(* IEC 61131-3 sources: trust-platform/tests/corpus, 4 files *)

(* ---- control_flow.st ---- *)
(* Test corpus: Control flow statements *)

PROGRAM TestControlFlow

VAR
    i, j, k : INT;
    condition : BOOL;
    state : INT;
    result : INT;
    sum : INT;
    arr : ARRAY[0..9] OF INT;
END_VAR

(* Simple IF *)
IF condition THEN
    result := 1;
END_IF

(* IF-ELSE *)
IF condition THEN
    result := 1;
ELSE
    result := 0;
END_IF

(* IF-ELSIF-ELSE *)
IF i < 0 THEN
    result := -1;
ELSIF i = 0 THEN
    result := 0;
ELSIF i > 0 AND i < 10 THEN
    result := 1;
ELSE
    result := 2;
END_IF

(* Nested IF *)
IF condition THEN
    IF i > 0 THEN
        result := 1;
    ELSE
        result := 2;
    END_IF
END_IF

(* Simple CASE *)
CASE state OF
    0: result := 0;
    1: result := 1;
    2: result := 2;
END_CASE

(* CASE with multiple labels *)
CASE state OF
    0, 1, 2:
        result := 0;
    3, 4, 5:
        result := 1;
    6..10:
        result := 2;
END_CASE

(* CASE with ELSE *)
CASE state OF
    0:
        result := 0;
    1:
        result := 1;
ELSE
    result := -1;
END_CASE

(* CASE with multiple statements *)
CASE state OF
    0:
        result := 0;
        condition := FALSE;
    1:
        result := 1;
        condition := TRUE;
END_CASE

(* Simple FOR *)
FOR i := 0 TO 9 DO
    arr[i] := i;
END_FOR

(* FOR with BY *)
FOR i := 0 TO 100 BY 10 DO
    sum := sum + i;
END_FOR

(* FOR counting down *)
FOR i := 10 TO 0 BY -1 DO
    arr[i] := i * 2;
END_FOR

(* Nested FOR *)
FOR i := 0 TO 9 DO
    FOR j := 0 TO 9 DO
        result := i * 10 + j;
    END_FOR
END_FOR

(* Simple WHILE *)
i := 0;
WHILE i < 10 DO
    sum := sum + i;
    i := i + 1;
END_WHILE

(* WHILE with complex condition *)
WHILE i < 10 AND NOT condition DO
    i := i + 1;
END_WHILE

(* Nested WHILE *)
i := 0;
WHILE i < 5 DO
    j := 0;
    WHILE j < 5 DO
        result := i * j;
        j := j + 1;
    END_WHILE
    i := i + 1;
END_WHILE

(* Simple REPEAT *)
i := 0;
REPEAT
    sum := sum + i;
    i := i + 1;
UNTIL i >= 10
END_REPEAT

(* REPEAT with complex condition *)
REPEAT
    i := i + 1;
    condition := i MOD 2 = 0;
UNTIL condition OR i > 100
END_REPEAT

(* EXIT from loop *)
FOR i := 0 TO 100 DO
    IF i > 50 THEN
        EXIT;
    END_IF
    sum := sum + i;
END_FOR

(* CONTINUE in loop *)
FOR i := 0 TO 9 DO
    IF i MOD 2 = 0 THEN
        CONTINUE;
    END_IF
    sum := sum + i;
END_FOR

(* EXIT from nested loop *)
FOR i := 0 TO 9 DO
    FOR j := 0 TO 9 DO
        IF i * j > 50 THEN
            EXIT;
        END_IF
    END_FOR
END_FOR

(* Empty statement *)
;

(* Multiple empty statements *)
;;

END_PROGRAM

(* Function with RETURN *)
FUNCTION CalcSum : INT
VAR_INPUT
    n : INT;
END_VAR
VAR
    i : INT;
    sum : INT;
END_VAR

IF n <= 0 THEN
    RETURN;
END_IF

FOR i := 1 TO n DO
    sum := sum + i;
END_FOR

CalcSum := sum;
END_FUNCTION

(* Function with early RETURN *)
FUNCTION FindIndex : INT
VAR_INPUT
    arr : ARRAY[0..9] OF INT;
    value : INT;
END_VAR
VAR
    i : INT;
END_VAR

FOR i := 0 TO 9 DO
    IF arr[i] = value THEN
        FindIndex := i;
        RETURN;
    END_IF
END_FOR

FindIndex := -1;
END_FUNCTION

(* Complex control flow *)
FUNCTION_BLOCK FB_StateMachine
VAR
    state : INT;
    counter : INT;
    done : BOOL;
END_VAR

CASE state OF
    0: (* Init *)
        counter := 0;
        state := 1;

    1: (* Process *)
        WHILE counter < 100 AND NOT done DO
            counter := counter + 1;
            IF counter MOD 10 = 0 THEN
                (* Check condition *)
                IF counter > 50 THEN
                    done := TRUE;
                    EXIT;
                END_IF
            END_IF
        END_WHILE

        IF done THEN
            state := 2;
        END_IF

    2: (* Done *)
        ; (* Empty - wait *)
END_CASE

END_FUNCTION_BLOCK

(* ---- declarations.st ---- *)
(* Test corpus: Variable declarations and modifiers *)

PROGRAM TestDeclarations

(* Basic variable block *)
VAR
    simpleVar : INT;
    multipleVars, anotherVar : BOOL;
    initialized : REAL := 3.14;
END_VAR

(* Input variables *)
VAR_INPUT
    inputBool : BOOL;
    inputInt : INT := 100;
END_VAR

(* Output variables *)
VAR_OUTPUT
    outputStatus : BOOL;
    outputValue : REAL;
END_VAR

(* In-out variables *)
VAR_IN_OUT
    inoutData : ARRAY[0..9] OF INT;
END_VAR

(* Temporary variables *)
VAR_TEMP
    tempCounter : INT;
    tempBuffer : STRING[80];
END_VAR

(* Constant variables *)
VAR CONSTANT
    PI : REAL := 3.14159;
    MAX_SIZE : INT := 1000;
END_VAR

(* Retain variables *)
VAR RETAIN
    persistentCounter : UDINT;
END_VAR

(* Non-retain variables *)
VAR NON_RETAIN
    volatileData : REAL;
END_VAR

(* Persistent variables *)
VAR PERSISTENT
    savedState : INT;
END_VAR

(* All elementary types *)
VAR
    boolVal : BOOL;
    sintVal : SINT;
    intVal : INT;
    dintVal : DINT;
    lintVal : LINT;
    usintVal : USINT;
    uintVal : UINT;
    udintVal : UDINT;
    ulintVal : ULINT;
    realVal : REAL;
    lrealVal : LREAL;
    byteVal : BYTE;
    wordVal : WORD;
    dwordVal : DWORD;
    lwordVal : LWORD;
    stringVal : STRING;
    stringFixed : STRING[100];
    wstringVal : WSTRING;
    timeVal : TIME;
    ltimeVal : LTIME;
    dateVal : DATE;
    todVal : TIME_OF_DAY;
    dtVal : DATE_AND_TIME;
END_VAR

END_PROGRAM

(* Global variables - must be in CONFIGURATION per IEC 61131-3 *)
CONFIGURATION GlobalConfig
VAR_GLOBAL
    GlobalCounter : UDINT;
    GlobalStatus : BOOL;
END_VAR

VAR_GLOBAL CONSTANT
    APP_VERSION : STRING := '1.0.0';
END_VAR
END_CONFIGURATION

(* External variables *)
PROGRAM TestExternal
VAR_EXTERNAL
    ExternalRef : REAL;
END_VAR
END_PROGRAM

(* Static variables in function block *)
FUNCTION_BLOCK FB_WithStatic
VAR_STAT
    callCount : UDINT;
END_VAR

callCount := callCount + 1;
END_FUNCTION_BLOCK

(* Type declarations *)
TYPE MyInt : INT; END_TYPE

TYPE MyRange : INT (0..100); END_TYPE

TYPE MyArray : ARRAY[0..9] OF INT; END_TYPE

TYPE MyArray2D : ARRAY[0..9, 0..9] OF REAL; END_TYPE

TYPE MyPointer : POINTER TO INT; END_TYPE

TYPE MyRef : REF_TO REAL; END_TYPE

TYPE MyString : STRING[255]; END_TYPE

TYPE MyStruct :
STRUCT
    field1 : INT;
    field2 : REAL;
    field3 : STRING[50];
END_STRUCT
END_TYPE

TYPE MyUnion :
UNION
    asInt : DINT;
    asReal : REAL;
    asBytes : ARRAY[0..3] OF BYTE;
END_UNION
END_TYPE

TYPE Color :
(
    Red := 0,
    Green := 1,
    Blue := 2
);
END_TYPE

(* Function with parameters *)
FUNCTION Add : INT
VAR_INPUT
    a : INT;
    b : INT;
END_VAR

Add := a + b;
END_FUNCTION

(* Function block with inheritance *)
FUNCTION_BLOCK FB_Child EXTENDS FB_Parent IMPLEMENTS I_Interface
VAR
    childVar : INT;
END_VAR
END_FUNCTION_BLOCK

(* Interface declaration *)
INTERFACE I_Counter
    METHOD Increment : INT
    END_METHOD

    METHOD Reset
    END_METHOD

    PROPERTY Count : INT
    END_PROPERTY
END_INTERFACE

(* Method with access modifiers *)
FUNCTION_BLOCK FB_AccessTest
VAR PUBLIC
    publicVar : INT;
END_VAR

VAR PRIVATE
    privateVar : INT;
END_VAR

PROTECTED METHOD ProtectedMethod
END_METHOD

PUBLIC METHOD PublicMethod
END_METHOD

PRIVATE METHOD PrivateMethod
END_METHOD
END_FUNCTION_BLOCK

(* Property with getter and setter *)
FUNCTION_BLOCK FB_PropertyTest
VAR
    _value : INT;
END_VAR

PROPERTY Value : INT
    GET
        Value := _value;
    END_GET
    SET
        _value := Value;
    END_SET
END_PROPERTY
END_FUNCTION_BLOCK

(* Namespace *)
NAMESPACE MyApp
    FUNCTION_BLOCK FB_Nested
    END_FUNCTION_BLOCK
END_NAMESPACE

(* ---- expressions.st ---- *)
(* Test corpus: Expressions and operator precedence *)

PROGRAM TestExpressions

VAR
    a, b, c, d : INT;
    x, y, z : REAL;
    p, q, r : BOOL;
    s1, s2 : STRING;
    arr : ARRAY[0..9] OF INT;
    ptr : POINTER TO INT;
    fb : FB_Test;
END_VAR

(* ============================================= *)
(* Arithmetic operators *)
(* ============================================= *)

(* Addition *)
a := 1 + 2;
a := b + c;
x := 1.0 + 2.5;

(* Subtraction *)
a := 5 - 3;
a := b - c;
x := 10.0 - 3.5;

(* Multiplication *)
a := 3 * 4;
a := b * c;
x := 2.0 * 3.14;

(* Division *)
a := 10 / 2;
x := 10.0 / 3.0;

(* Modulo *)
a := 10 MOD 3;
a := b MOD c;

(* Exponentiation - right associative *)
x := 2.0 ** 3.0;
x := 2.0 ** 3.0 ** 2.0;  (* = 2^(3^2) = 2^9 = 512 *)

(* Unary operators *)
a := -b;
a := +c;
x := -3.14;

(* ============================================= *)
(* Comparison operators *)
(* ============================================= *)

p := a = b;
p := a <> b;
p := a < b;
p := a <= b;
p := a > b;
p := a >= b;

(* String comparison *)
p := s1 = s2;
p := s1 < s2;

(* ============================================= *)
(* Logical operators *)
(* ============================================= *)

(* AND *)
p := q AND r;
p := q & r;

(* OR *)
p := q OR r;

(* XOR *)
p := q XOR r;

(* NOT *)
p := NOT q;

(* ============================================= *)
(* Bitwise operators *)
(* ============================================= *)

a := b AND c;
a := b OR c;
a := b XOR c;
a := NOT b;

(* ============================================= *)
(* Operator precedence tests *)
(* ============================================= *)

(* Precedence: * before + *)
a := 1 + 2 * 3;         (* = 1 + 6 = 7 *)
a := (1 + 2) * 3;       (* = 3 * 3 = 9 *)

(* Precedence: AND before OR *)
p := TRUE OR FALSE AND FALSE;     (* = TRUE OR FALSE = TRUE *)
p := (TRUE OR FALSE) AND FALSE;   (* = TRUE AND FALSE = FALSE *)

(* Precedence: comparison before logical *)
p := a < b AND c > d;   (* = (a < b) AND (c > d) *)

(* Precedence: arithmetic before comparison *)
p := a + b < c + d;     (* = (a + b) < (c + d) *)

(* Precedence: NOT has highest priority *)
p := NOT q AND r;       (* = (NOT q) AND r *)
p := NOT (q AND r);     (* = NOT (q AND r) *)

(* Complex precedence *)
a := 1 + 2 * 3 - 4 / 2;     (* = 1 + 6 - 2 = 5 *)
p := a > b OR c < d AND NOT r;  (* = (a > b) OR ((c < d) AND (NOT r)) *)

(* Power is right associative *)
x := 2.0 ** 2.0 ** 3.0;     (* = 2^(2^3) = 2^8 = 256 *)

(* ============================================= *)
(* Parenthesized expressions *)
(* ============================================= *)

a := (b);
a := ((b));
a := (b + c);
a := (b + c) * d;
a := ((b + c) * (d - a));

(* ============================================= *)
(* Function calls *)
(* ============================================= *)

x := SIN(3.14);
x := ABS(-42);
a := MAX(b, c);
x := SQRT(y);

(* Nested function calls *)
x := SIN(COS(3.14));
x := ABS(MIN(a, b));

(* Function call in expression *)
x := 2.0 * SIN(y) + 1.0;

(* Named parameters *)
(* result := MyFunc(param1 := 10, param2 := 20); *)

(* ============================================= *)
(* Array indexing *)
(* ============================================= *)

a := arr[0];
a := arr[b];
a := arr[b + 1];
a := arr[b * 2 + c];

(* Multi-dimensional *)
(* a := matrix[i, j]; *)
(* a := matrix[i][j]; *)

(* ============================================= *)
(* Field access *)
(* ============================================= *)

a := fb.value;
x := fb.data.x;
a := fb.nested.deep.value;

(* Method call *)
a := fb.GetValue();
fb.SetValue(10);

(* ============================================= *)
(* Pointer operations *)
(* ============================================= *)

(* Dereference *)
a := ptr^;

(* Address-of *)
ptr := ADR(a);

(* SIZEOF *)
a := SIZEOF(INT);
a := SIZEOF(arr);
a := SIZEOF(fb);

(* ============================================= *)
(* Special expressions *)
(* ============================================= *)

(* THIS and SUPER *)
(* a := THIS.value; *)
(* a := SUPER.GetValue(); *)

(* Direct addresses *)
(* a := %IW10; *)
(* p := %IX0.0; *)

(* Typed literals in expressions *)
a := INT#42 + INT#10;
x := REAL#3.14 * REAL#2.0;

(* ============================================= *)
(* Complex expressions *)
(* ============================================= *)

(* Combined arithmetic and logic *)
p := (a + b > c) AND (d - a < 10) OR NOT q;

(* Expression with function call and array *)
a := arr[MAX(b, c)] + ABS(d);

(* Expression with field access *)
x := fb.value * SIN(fb.angle);

(* Very complex expression *)
x := ((a + b) * SIN(c / d)) / (SQRT(y ** 2.0 + z ** 2.0) + 1.0);

END_PROGRAM

(* Function block for testing *)
FUNCTION_BLOCK FB_Test
VAR
    value : INT;
    angle : REAL;
    data : ST_Data;
    nested : FB_Nested;
END_VAR

METHOD GetValue : INT
    GetValue := value;
END_METHOD

METHOD SetValue
VAR_INPUT
    newValue : INT;
END_VAR
    value := newValue;
END_METHOD
END_FUNCTION_BLOCK

FUNCTION_BLOCK FB_Nested
VAR
    deep : ST_Deep;
END_VAR
END_FUNCTION_BLOCK

TYPE ST_Data :
STRUCT
    x : REAL;
    y : REAL;
END_STRUCT
END_TYPE

TYPE ST_Deep :
STRUCT
    value : INT;
END_STRUCT
END_TYPE

(* Test expression edge cases *)
FUNCTION TestEdgeCases : BOOL
VAR
    a : INT;
    x : REAL;
    p : BOOL;
END_VAR

(* Double negation *)
a := --5;
a := -(-a);
x := --3.14;

(* NOT NOT *)
p := NOT NOT TRUE;
p := NOT NOT p;

(* Chained comparisons need explicit grouping *)
p := (a < 5) AND (5 < 10);

(* Very deep nesting *)
a := ((((((1 + 2) * 3) - 4) / 5) MOD 6) + 7);

TestEdgeCases := TRUE;
END_FUNCTION

(* ---- literals.st ---- *)
(* Test corpus: All literal types *)

PROGRAM TestLiterals

VAR
    (* Integer literals *)
    intDec : INT := 123;
    intNeg : INT := -456;
    intZero : INT := 0;
    intWithUnder : DINT := 1_000_000;

    (* Hexadecimal literals *)
    intHex : DWORD := 16#FF;
    intHexLower : DWORD := 16#ff;
    intHexMixed : DWORD := 16#DeAdBeEf;
    intHexUnder : DWORD := 16#DEAD_BEEF;

    (* Binary literals *)
    intBin : BYTE := 2#10101010;
    intBinUnder : WORD := 2#1111_0000_1111_0000;

    (* Octal literals *)
    intOct : INT := 8#77;
    intOctUnder : INT := 8#7_7_7;

    (* Real literals *)
    realSimple : REAL := 3.14;
    realNeg : REAL := -2.718;
    realZero : REAL := 0.0;
    realSmall : REAL := 0.001;
    realWithUnder : LREAL := 1_000.000_001;

    (* Scientific notation *)
    realSci1 : LREAL := 1.0E10;
    realSci2 : LREAL := 2.5e-3;
    realSci3 : LREAL := 6.022E+23;
    realSciNeg : LREAL := -1.6E-19;

    (* Boolean literals *)
    boolTrue : BOOL := TRUE;
    boolFalse : BOOL := FALSE;
    boolTrueLower : BOOL := true;
    boolFalseLower : BOOL := false;

    (* String literals - single quote *)
    strEmpty : STRING := '';
    strSimple : STRING := 'Hello, World!';
    strWithEscape : STRING := 'Line1$NLine2';
    strWithQuote : STRING := 'It$'s working';
    strPath : STRING := 'C:\Program Files\App';

    (* Wide string literals - double quote *)
    wstrEmpty : WSTRING := "";
    wstrSimple : WSTRING := "Wide string";
    wstrUnicode : WSTRING := "日本語";

    (* Time literals *)
    timeSimple : TIME := T#1s;
    timeLong : TIME := TIME#1h30m45s;
    timeMs : TIME := T#100ms;
    timeComplex : TIME := T#1d2h3m4s5ms;
    timeUnder : TIME := T#1000ms;
    ltimeVal : LTIME := LTIME#1h;

    (* Date literals *)
    dateSimple : DATE := D#2024-01-15;
    dateFull : DATE := DATE#2024-12-31;

    (* Time of day literals *)
    todSimple : TIME_OF_DAY := TOD#12:30:00;
    todFull : TIME_OF_DAY := TIME_OF_DAY#23:59:59.999;
    todMidnight : TIME_OF_DAY := TOD#00:00:00;

    (* Date and time literals *)
    dtSimple : DATE_AND_TIME := DT#2024-01-15-12:30:00;
    dtFull : DATE_AND_TIME := DATE_AND_TIME#2024-12-31-23:59:59;
END_VAR

VAR
    (* Typed literals *)
    typedInt : INT := INT#42;
    typedDint : DINT := DINT#1000000;
    typedReal : REAL := REAL#3.14;
    typedBool : BOOL := BOOL#TRUE;
    typedByte : BYTE := BYTE#16#FF;
    typedWord : WORD := WORD#2#1010101010101010;
    typedLreal : LREAL := LREAL#1.0E-10;

    (* Typed literals with type prefix *)
    hexTyped : DWORD := DWORD#16#DEADBEEF;
    binTyped : BYTE := BYTE#2#11110000;

    (* Enum typed literals - common pattern *)
    (* enumVal : MyEnum := MyEnum#Value1; *)
END_VAR

VAR CONSTANT
    (* Constants with various literal types *)
    CONST_PI : LREAL := 3.14159265358979;
    CONST_E : LREAL := 2.71828182845905;
    CONST_MAX_INT : DINT := 2147483647;
    CONST_MIN_INT : DINT := -2147483648;
    CONST_HEX : DWORD := 16#FFFFFFFF;
    CONST_TIMEOUT : TIME := T#30s;
    CONST_MSG : STRING := 'Constant message';
END_VAR

END_PROGRAM

(* Test literals in expressions *)
FUNCTION TestLiteralExpressions : BOOL
VAR
    result : REAL;
    flag : BOOL;
    text : STRING;
END_VAR

(* Literals in arithmetic *)
result := 10 + 20;
result := 3.14 * 2.0;
result := 16#FF + 1;
result := 2#1010 AND 2#1100;

(* Literals in comparisons *)
flag := 100 > 50;
flag := 3.14 < 4.0;
flag := 'abc' < 'abd';

(* Literals in function calls *)
result := SIN(3.14159);
result := ABS(-42);

(* Time arithmetic *)
(* delay := T#1s + T#500ms; *)

(* Literals in array access *)
(* arr[0] := 1; *)
(* arr[16#0A] := 10; *)

TestLiteralExpressions := TRUE;
END_FUNCTION

(* Test edge cases *)
PROGRAM TestLiteralEdgeCases
VAR
    (* Very large numbers *)
    bigInt : LINT := 9223372036854775807;
    bigReal : LREAL := 1.7976931348623157E+308;

    (* Very small numbers *)
    smallReal : LREAL := 2.2250738585072014E-308;

    (* Zero variants *)
    zeroInt : INT := 0;
    zeroReal : REAL := 0.0;
    zeroHex : DWORD := 16#0;
    zeroBin : BYTE := 2#0;

    (* Long strings *)
    longStr : STRING[255] := 'This is a very long string that contains many characters and is used to test the parser handling of long string literals in the source code.';
END_VAR
END_PROGRAM
